# EPICS substitutions: db/Beckhoff_7XXX/ecmcEP7211-0034_OPT_csp.substitutions
file "ecmcEL72XX_DRV_CSP.template"
{
  pattern {CH_ID}
          {01   }
}
